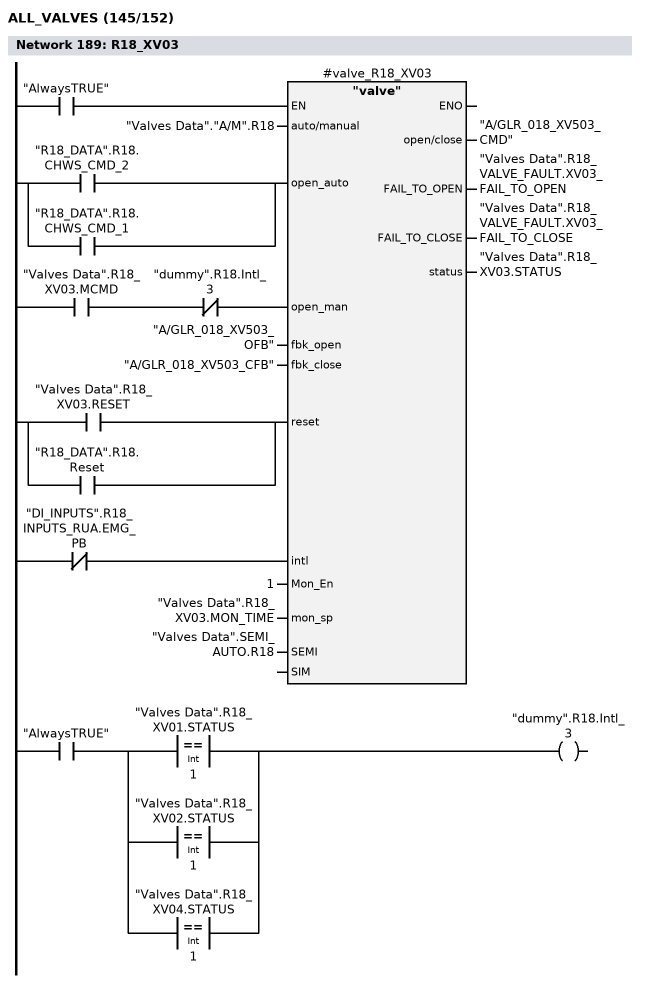
   RUNG wire#powerrail
      Contact( "AlwaysTRUE" )
      #valve_R18_XV03(open_auto := wire#w1, open_man := wire#w2, reset := wire#w3, intl := wire#w4, "auto/manual" := "Valves Data"."A/M".R18, fbk_open := "A/GLR_018_XV503_OFB", fbk_close := "A/GLR_018_XV503_CFB", Mon_En := 1, mon_sp := "Valves Data".R18_XV03.MON_TIME, SEMI := "Valves Data".SEMI_AUTO.R18, SIM :=, "open/close" => "A/GLR_018_XV503_CMD", FAIL_TO_OPEN => "Valves Data".R18_VALVE_FAULT.XV03_FAIL_TO_OPEN, FAIL_TO_CLOSE => "Valves Data".R18_VALVE_FAULT.XV03_FAIL_TO_CLOSE, status => "Valves Data".R18_XV03.STATUS)
   END_RUNG
   RUNG wire#powerrail
      Contact( "R18_DATA".R18.CHWS_CMD_2 )
   END_RUNG wire#w1
   RUNG wire#powerrail
      Contact( "R18_DATA".R18.CHWS_CMD_1 )
   END_RUNG wire#w1
   RUNG wire#powerrail
      Contact( "Valves Data".R18_XV03.MCMD )
      I_Contact( "dummy".R18.Intl_3 )
   END_RUNG wire#w2
   RUNG wire#powerrail
      Contact( "Valves Data".R18_XV03.RESET )
   END_RUNG wire#w3
   RUNG wire#powerrail
      Contact( "R18_DATA".R18.Reset )
   END_RUNG wire#w3
   RUNG wire#powerrail
      I_Contact( "DI_INPUTS".R18_INPUTS_RUA.EMG_PB )
   END_RUNG wire#w4
   RUNG wire#powerrail
      Contact( "AlwaysTRUE" )
      wire#w5
      { S7_Templates := "SrcType := Int" } EQ_Contact(in1 := "Valves Data".R18_XV01.STATUS, in2 := 1)
      wire#w6
      Coil( "dummy".R18.Intl_3 )
   END_RUNG
   RUNG wire#w5
      { S7_Templates := "SrcType := Int" } EQ_Contact(in1 := "Valves Data".R18_XV02.STATUS, in2 := 1)
   END_RUNG wire#w6
   RUNG wire#w5
      { S7_Templates := "SrcType := Int" } EQ_Contact(in1 := "Valves Data".R18_XV04.STATUS, in2 := 1)
   END_RUNG wire#w6
   // the same network as SCL:
   IF "AlwaysTRUE" THEN
       #valve_R18_XV03("auto/manual" := "Valves Data"."A/M".R18,   // "valve"
                       open_auto := "R18_DATA".R18.CHWS_CMD_2 OR "R18_DATA".R18.CHWS_CMD_1,
                       open_man := "Valves Data".R18_XV03.MCMD AND NOT "dummy".R18.Intl_3,
                       fbk_open := "A/GLR_018_XV503_OFB",
                       fbk_close := "A/GLR_018_XV503_CFB",
                       reset := "Valves Data".R18_XV03.RESET OR "R18_DATA".R18.Reset,
                       intl := NOT "DI_INPUTS".R18_INPUTS_RUA.EMG_PB,
                       Mon_En := 1,
                       mon_sp := "Valves Data".R18_XV03.MON_TIME,
                       SEMI := "Valves Data".SEMI_AUTO.R18,
                       "open/close" => "A/GLR_018_XV503_CMD",
                       FAIL_TO_OPEN => "Valves Data".R18_VALVE_FAULT.XV03_FAIL_TO_OPEN,
                       FAIL_TO_CLOSE => "Valves Data".R18_VALVE_FAULT.XV03_FAIL_TO_CLOSE,
                       status => "Valves Data".R18_XV03.STATUS);
   END_IF;
   "dummy".R18.Intl_3 := "AlwaysTRUE" AND (("Valves Data".R18_XV01.STATUS = 1) OR ("Valves Data".R18_XV02.STATUS = 1) OR ("Valves Data".R18_XV04.STATUS = 1));
END_REGION

REGION Network 190: R18_XV04
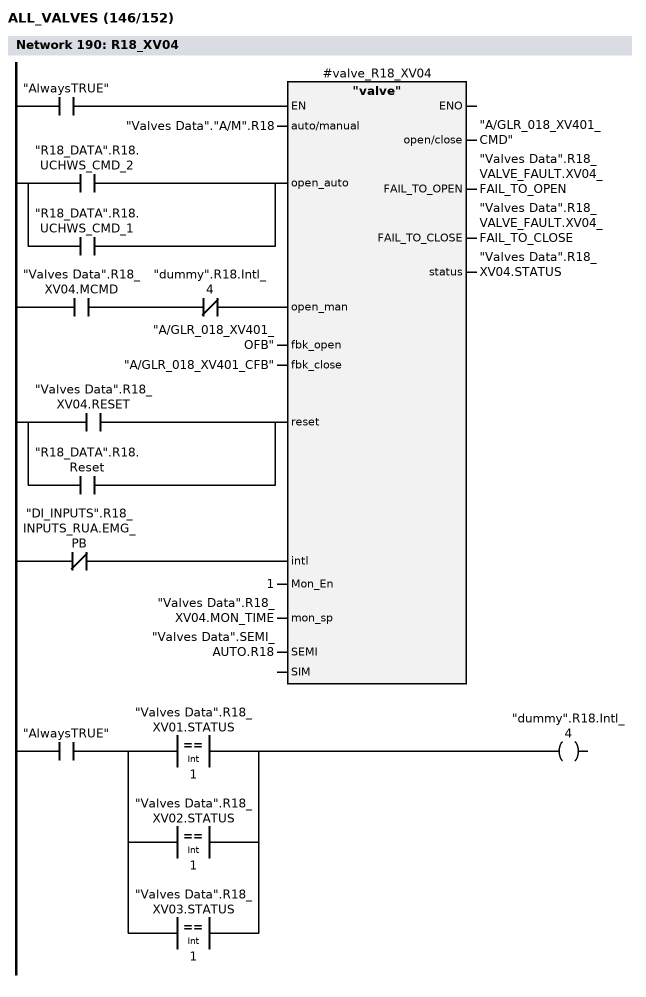
   RUNG wire#powerrail
      Contact( "AlwaysTRUE" )
      #valve_R18_XV04(open_auto := wire#w1, open_man := wire#w2, reset := wire#w3, intl := wire#w4, "auto/manual" := "Valves Data"."A/M".R18, fbk_open := "A/GLR_018_XV401_OFB", fbk_close := "A/GLR_018_XV401_CFB", Mon_En := 1, mon_sp := "Valves Data".R18_XV04.MON_TIME, SEMI := "Valves Data".SEMI_AUTO.R18, SIM :=, "open/close" => "A/GLR_018_XV401_CMD", FAIL_TO_OPEN => "Valves Data".R18_VALVE_FAULT.XV04_FAIL_TO_OPEN, FAIL_TO_CLOSE => "Valves Data".R18_VALVE_FAULT.XV04_FAIL_TO_CLOSE, status => "Valves Data".R18_XV04.STATUS)
   END_RUNG
   RUNG wire#powerrail
      Contact( "R18_DATA".R18.UCHWS_CMD_2 )
   END_RUNG wire#w1
   RUNG wire#powerrail
      Contact( "R18_DATA".R18.UCHWS_CMD_1 )
   END_RUNG wire#w1
   RUNG wire#powerrail
      Contact( "Valves Data".R18_XV04.MCMD )
      I_Contact( "dummy".R18.Intl_4 )
   END_RUNG wire#w2
   RUNG wire#powerrail
      Contact( "Valves Data".R18_XV04.RESET )
   END_RUNG wire#w3
   RUNG wire#powerrail
      Contact( "R18_DATA".R18.Reset )
   END_RUNG wire#w3
   RUNG wire#powerrail
      I_Contact( "DI_INPUTS".R18_INPUTS_RUA.EMG_PB )
   END_RUNG wire#w4
   RUNG wire#powerrail
      Contact( "AlwaysTRUE" )
      wire#w5
      { S7_Templates := "SrcType := Int" } EQ_Contact(in1 := "Valves Data".R18_XV01.STATUS, in2 := 1)
      wire#w6
      Coil( "dummy".R18.Intl_4 )
   END_RUNG
   RUNG wire#w5
      { S7_Templates := "SrcType := Int" } EQ_Contact(in1 := "Valves Data".R18_XV02.STATUS, in2 := 1)
   END_RUNG wire#w6
   RUNG wire#w5
      { S7_Templates := "SrcType := Int" } EQ_Contact(in1 := "Valves Data".R18_XV03.STATUS, in2 := 1)
   END_RUNG wire#w6
   // the same network as SCL:
   IF "AlwaysTRUE" THEN
       #valve_R18_XV04("auto/manual" := "Valves Data"."A/M".R18,   // "valve"
                       open_auto := "R18_DATA".R18.UCHWS_CMD_2 OR "R18_DATA".R18.UCHWS_CMD_1,
                       open_man := "Valves Data".R18_XV04.MCMD AND NOT "dummy".R18.Intl_4,
                       fbk_open := "A/GLR_018_XV401_OFB",
                       fbk_close := "A/GLR_018_XV401_CFB",
                       reset := "Valves Data".R18_XV04.RESET OR "R18_DATA".R18.Reset,
                       intl := NOT "DI_INPUTS".R18_INPUTS_RUA.EMG_PB,
                       Mon_En := 1,
                       mon_sp := "Valves Data".R18_XV04.MON_TIME,
                       SEMI := "Valves Data".SEMI_AUTO.R18,
                       "open/close" => "A/GLR_018_XV401_CMD",
                       FAIL_TO_OPEN => "Valves Data".R18_VALVE_FAULT.XV04_FAIL_TO_OPEN,
                       FAIL_TO_CLOSE => "Valves Data".R18_VALVE_FAULT.XV04_FAIL_TO_CLOSE,
                       status => "Valves Data".R18_XV04.STATUS);
   END_IF;
   "dummy".R18.Intl_4 := "AlwaysTRUE" AND (("Valves Data".R18_XV01.STATUS = 1) OR ("Valves Data".R18_XV02.STATUS = 1) OR ("Valves Data".R18_XV03.STATUS = 1));
END_REGION

REGION Network 191: R18_XV05
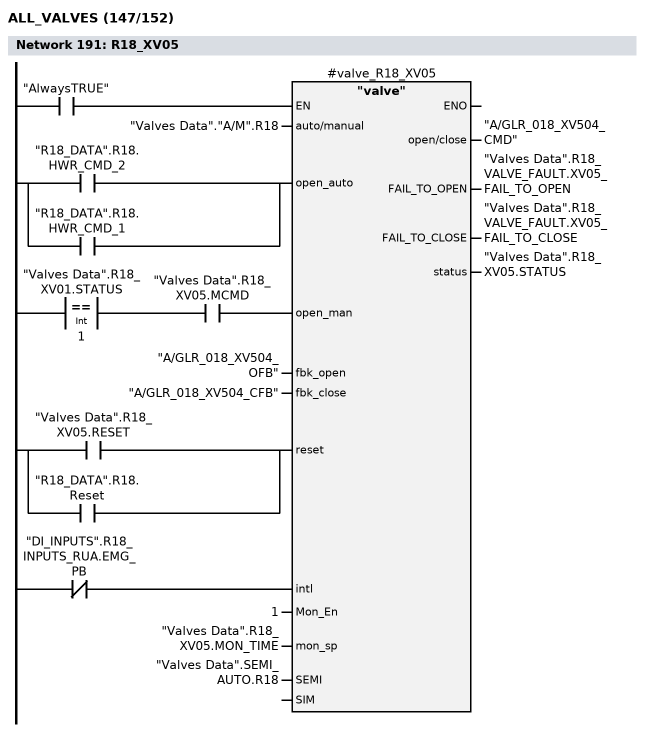
   RUNG wire#powerrail
      Contact( "AlwaysTRUE" )
      #valve_R18_XV05(open_auto := wire#w1, open_man := wire#w2, reset := wire#w3, intl := wire#w4, "auto/manual" := "Valves Data"."A/M".R18, fbk_open := "A/GLR_018_XV504_OFB", fbk_close := "A/GLR_018_XV504_CFB", Mon_En := 1, mon_sp := "Valves Data".R18_XV05.MON_TIME, SEMI := "Valves Data".SEMI_AUTO.R18, SIM :=, "open/close" => "A/GLR_018_XV504_CMD", FAIL_TO_OPEN => "Valves Data".R18_VALVE_FAULT.XV05_FAIL_TO_OPEN, FAIL_TO_CLOSE => "Valves Data".R18_VALVE_FAULT.XV05_FAIL_TO_CLOSE, status => "Valves Data".R18_XV05.STATUS)
   END_RUNG
   RUNG wire#powerrail
      Contact( "R18_DATA".R18.HWR_CMD_2 )
   END_RUNG wire#w1
   RUNG wire#powerrail
      Contact( "R18_DATA".R18.HWR_CMD_1 )
   END_RUNG wire#w1
   RUNG wire#powerrail
      { S7_Templates := "SrcType := Int" } EQ_Contact(in1 := "Valves Data".R18_XV01.STATUS, in2 := 1)
      Contact( "Valves Data".R18_XV05.MCMD )
   END_RUNG wire#w2
   RUNG wire#powerrail
      Contact( "Valves Data".R18_XV05.RESET )
   END_RUNG wire#w3
   RUNG wire#powerrail
      Contact( "R18_DATA".R18.Reset )
   END_RUNG wire#w3
   RUNG wire#powerrail
      I_Contact( "DI_INPUTS".R18_INPUTS_RUA.EMG_PB )
   END_RUNG wire#w4
   // the same network as SCL:
   IF "AlwaysTRUE" THEN
       #valve_R18_XV05("auto/manual" := "Valves Data"."A/M".R18,   // "valve"
                       open_auto := "R18_DATA".R18.HWR_CMD_2 OR "R18_DATA".R18.HWR_CMD_1,
                       open_man := ("Valves Data".R18_XV01.STATUS = 1) AND "Valves Data".R18_XV05.MCMD,
                       fbk_open := "A/GLR_018_XV504_OFB",
                       fbk_close := "A/GLR_018_XV504_CFB",
                       reset := "Valves Data".R18_XV05.RESET OR "R18_DATA".R18.Reset,
                       intl := NOT "DI_INPUTS".R18_INPUTS_RUA.EMG_PB,
                       Mon_En := 1,
                       mon_sp := "Valves Data".R18_XV05.MON_TIME,
                       SEMI := "Valves Data".SEMI_AUTO.R18,
                       "open/close" => "A/GLR_018_XV504_CMD",
                       FAIL_TO_OPEN => "Valves Data".R18_VALVE_FAULT.XV05_FAIL_TO_OPEN,
                       FAIL_TO_CLOSE => "Valves Data".R18_VALVE_FAULT.XV05_FAIL_TO_CLOSE,
                       status => "Valves Data".R18_XV05.STATUS);
   END_IF;
END_REGION

REGION Network 192: R18_XV06
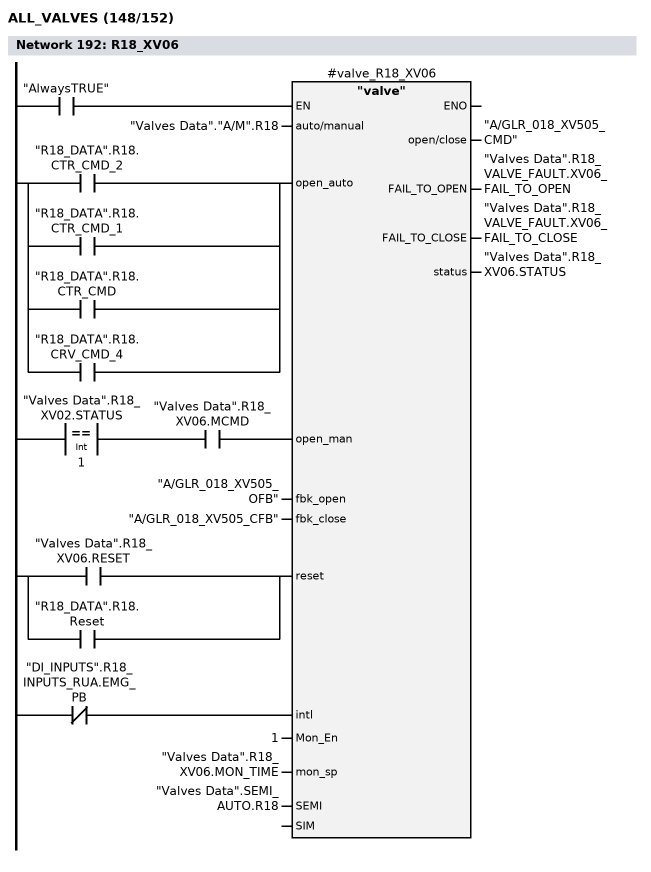
   RUNG wire#powerrail
      Contact( "AlwaysTRUE" )
      #valve_R18_XV06(open_auto := wire#w1, open_man := wire#w2, reset := wire#w3, intl := wire#w4, "auto/manual" := "Valves Data"."A/M".R18, fbk_open := "A/GLR_018_XV505_OFB", fbk_close := "A/GLR_018_XV505_CFB", Mon_En := 1, mon_sp := "Valves Data".R18_XV06.MON_TIME, SEMI := "Valves Data".SEMI_AUTO.R18, SIM :=, "open/close" => "A/GLR_018_XV505_CMD", FAIL_TO_OPEN => "Valves Data".R18_VALVE_FAULT.XV06_FAIL_TO_OPEN, FAIL_TO_CLOSE => "Valves Data".R18_VALVE_FAULT.XV06_FAIL_TO_CLOSE, status => "Valves Data".R18_XV06.STATUS)
   END_RUNG
   RUNG wire#powerrail
      Contact( "R18_DATA".R18.CTR_CMD_2 )
   END_RUNG wire#w1
   RUNG wire#powerrail
      Contact( "R18_DATA".R18.CTR_CMD_1 )
   END_RUNG wire#w1
   RUNG wire#powerrail
      Contact( "R18_DATA".R18.CTR_CMD )
   END_RUNG wire#w1
   RUNG wire#powerrail
      Contact( "R18_DATA".R18.CRV_CMD_4 )
   END_RUNG wire#w1
   RUNG wire#powerrail
      { S7_Templates := "SrcType := Int" } EQ_Contact(in1 := "Valves Data".R18_XV02.STATUS, in2 := 1)
      Contact( "Valves Data".R18_XV06.MCMD )
   END_RUNG wire#w2
   RUNG wire#powerrail
      Contact( "Valves Data".R18_XV06.RESET )
   END_RUNG wire#w3
   RUNG wire#powerrail
      Contact( "R18_DATA".R18.Reset )
   END_RUNG wire#w3
   RUNG wire#powerrail
      I_Contact( "DI_INPUTS".R18_INPUTS_RUA.EMG_PB )
   END_RUNG wire#w4
   // the same network as SCL:
   IF "AlwaysTRUE" THEN
       #valve_R18_XV06("auto/manual" := "Valves Data"."A/M".R18,   // "valve"
                       open_auto := "R18_DATA".R18.CTR_CMD_2 OR "R18_DATA".R18.CTR_CMD_1 OR "R18_DATA".R18.CTR_CMD OR "R18_DATA".R18.CRV_CMD_4,
                       open_man := ("Valves Data".R18_XV02.STATUS = 1) AND "Valves Data".R18_XV06.MCMD,
                       fbk_open := "A/GLR_018_XV505_OFB",
                       fbk_close := "A/GLR_018_XV505_CFB",
                       reset := "Valves Data".R18_XV06.RESET OR "R18_DATA".R18.Reset,
                       intl := NOT "DI_INPUTS".R18_INPUTS_RUA.EMG_PB,
                       Mon_En := 1,
                       mon_sp := "Valves Data".R18_XV06.MON_TIME,
                       SEMI := "Valves Data".SEMI_AUTO.R18,
                       "open/close" => "A/GLR_018_XV505_CMD",
                       FAIL_TO_OPEN => "Valves Data".R18_VALVE_FAULT.XV06_FAIL_TO_OPEN,
                       FAIL_TO_CLOSE => "Valves Data".R18_VALVE_FAULT.XV06_FAIL_TO_CLOSE,
                       status => "Valves Data".R18_XV06.STATUS);
   END_IF;
END_REGION

REGION Network 193: R18_XV07
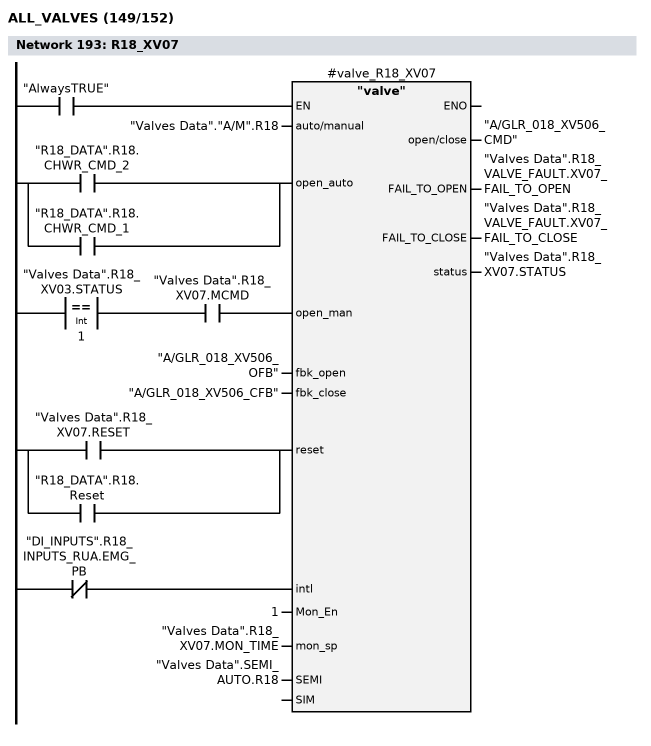
   RUNG wire#powerrail
      Contact( "AlwaysTRUE" )
      #valve_R18_XV07(open_auto := wire#w1, open_man := wire#w2, reset := wire#w3, intl := wire#w4, "auto/manual" := "Valves Data"."A/M".R18, fbk_open := "A/GLR_018_XV506_OFB", fbk_close := "A/GLR_018_XV506_CFB", Mon_En := 1, mon_sp := "Valves Data".R18_XV07.MON_TIME, SEMI := "Valves Data".SEMI_AUTO.R18, SIM :=, "open/close" => "A/GLR_018_XV506_CMD", FAIL_TO_OPEN => "Valves Data".R18_VALVE_FAULT.XV07_FAIL_TO_OPEN, FAIL_TO_CLOSE => "Valves Data".R18_VALVE_FAULT.XV07_FAIL_TO_CLOSE, status => "Valves Data".R18_XV07.STATUS)
   END_RUNG
   RUNG wire#powerrail
      Contact( "R18_DATA".R18.CHWR_CMD_2 )
   END_RUNG wire#w1
   RUNG wire#powerrail
      Contact( "R18_DATA".R18.CHWR_CMD_1 )
   END_RUNG wire#w1
   RUNG wire#powerrail
      { S7_Templates := "SrcType := Int" } EQ_Contact(in1 := "Valves Data".R18_XV03.STATUS, in2 := 1)
      Contact( "Valves Data".R18_XV07.MCMD )
   END_RUNG wire#w2
   RUNG wire#powerrail
      Contact( "Valves Data".R18_XV07.RESET )
   END_RUNG wire#w3
   RUNG wire#powerrail
      Contact( "R18_DATA".R18.Reset )
   END_RUNG wire#w3
   RUNG wire#powerrail
      I_Contact( "DI_INPUTS".R18_INPUTS_RUA.EMG_PB )
   END_RUNG wire#w4
   // the same network as SCL:
   IF "AlwaysTRUE" THEN
       #valve_R18_XV07("auto/manual" := "Valves Data"."A/M".R18,   // "valve"
                       open_auto := "R18_DATA".R18.CHWR_CMD_2 OR "R18_DATA".R18.CHWR_CMD_1,
                       open_man := ("Valves Data".R18_XV03.STATUS = 1) AND "Valves Data".R18_XV07.MCMD,
                       fbk_open := "A/GLR_018_XV506_OFB",
                       fbk_close := "A/GLR_018_XV506_CFB",
                       reset := "Valves Data".R18_XV07.RESET OR "R18_DATA".R18.Reset,
                       intl := NOT "DI_INPUTS".R18_INPUTS_RUA.EMG_PB,
                       Mon_En := 1,
                       mon_sp := "Valves Data".R18_XV07.MON_TIME,
                       SEMI := "Valves Data".SEMI_AUTO.R18,
                       "open/close" => "A/GLR_018_XV506_CMD",
                       FAIL_TO_OPEN => "Valves Data".R18_VALVE_FAULT.XV07_FAIL_TO_OPEN,
                       FAIL_TO_CLOSE => "Valves Data".R18_VALVE_FAULT.XV07_FAIL_TO_CLOSE,
                       status => "Valves Data".R18_XV07.STATUS);
   END_IF;
END_REGION

REGION Network 194: R18_XV08
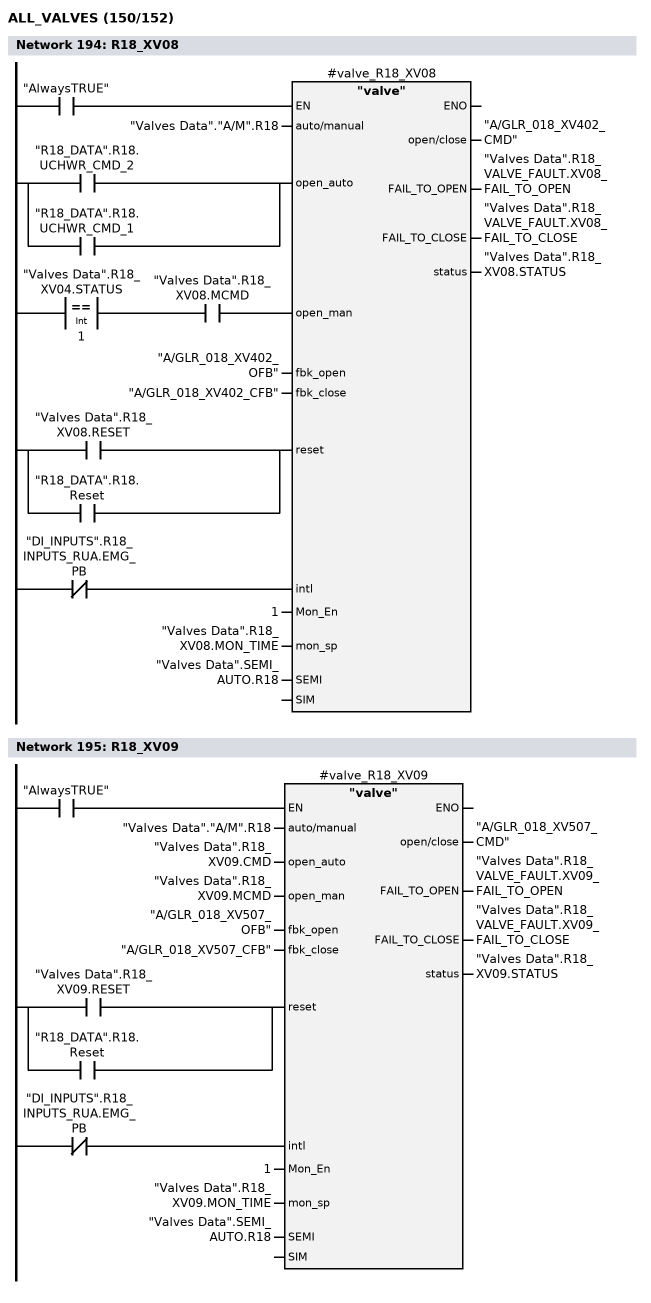
   RUNG wire#powerrail
      Contact( "AlwaysTRUE" )
      #valve_R18_XV08(open_auto := wire#w1, open_man := wire#w2, reset := wire#w3, intl := wire#w4, "auto/manual" := "Valves Data"."A/M".R18, fbk_open := "A/GLR_018_XV402_OFB", fbk_close := "A/GLR_018_XV402_CFB", Mon_En := 1, mon_sp := "Valves Data".R18_XV08.MON_TIME, SEMI := "Valves Data".SEMI_AUTO.R18, SIM :=, "open/close" => "A/GLR_018_XV402_CMD", FAIL_TO_OPEN => "Valves Data".R18_VALVE_FAULT.XV08_FAIL_TO_OPEN, FAIL_TO_CLOSE => "Valves Data".R18_VALVE_FAULT.XV08_FAIL_TO_CLOSE, status => "Valves Data".R18_XV08.STATUS)
   END_RUNG
   RUNG wire#powerrail
      Contact( "R18_DATA".R18.UCHWR_CMD_2 )
   END_RUNG wire#w1
   RUNG wire#powerrail
      Contact( "R18_DATA".R18.UCHWR_CMD_1 )
   END_RUNG wire#w1
   RUNG wire#powerrail
      { S7_Templates := "SrcType := Int" } EQ_Contact(in1 := "Valves Data".R18_XV04.STATUS, in2 := 1)
      Contact( "Valves Data".R18_XV08.MCMD )
   END_RUNG wire#w2
   RUNG wire#powerrail
      Contact( "Valves Data".R18_XV08.RESET )
   END_RUNG wire#w3
   RUNG wire#powerrail
      Contact( "R18_DATA".R18.Reset )
   END_RUNG wire#w3
   RUNG wire#powerrail
      I_Contact( "DI_INPUTS".R18_INPUTS_RUA.EMG_PB )
   END_RUNG wire#w4
   // the same network as SCL:
   IF "AlwaysTRUE" THEN
       #valve_R18_XV08("auto/manual" := "Valves Data"."A/M".R18,   // "valve"
                       open_auto := "R18_DATA".R18.UCHWR_CMD_2 OR "R18_DATA".R18.UCHWR_CMD_1,
                       open_man := ("Valves Data".R18_XV04.STATUS = 1) AND "Valves Data".R18_XV08.MCMD,
                       fbk_open := "A/GLR_018_XV402_OFB",
                       fbk_close := "A/GLR_018_XV402_CFB",
                       reset := "Valves Data".R18_XV08.RESET OR "R18_DATA".R18.Reset,
                       intl := NOT "DI_INPUTS".R18_INPUTS_RUA.EMG_PB,
                       Mon_En := 1,
                       mon_sp := "Valves Data".R18_XV08.MON_TIME,
                       SEMI := "Valves Data".SEMI_AUTO.R18,
                       "open/close" => "A/GLR_018_XV402_CMD",
                       FAIL_TO_OPEN => "Valves Data".R18_VALVE_FAULT.XV08_FAIL_TO_OPEN,
                       FAIL_TO_CLOSE => "Valves Data".R18_VALVE_FAULT.XV08_FAIL_TO_CLOSE,
                       status => "Valves Data".R18_XV08.STATUS);
   END_IF;
END_REGION

REGION Network 195: R18_XV09
   RUNG wire#powerrail
      Contact( "AlwaysTRUE" )
      #valve_R18_XV09(reset := wire#w1, intl := wire#w2, "auto/manual" := "Valves Data"."A/M".R18, open_auto := "Valves Data".R18_XV09.CMD, open_man := "Valves Data".R18_XV09.MCMD, fbk_open := "A/GLR_018_XV507_OFB", fbk_close := "A/GLR_018_XV507_CFB", Mon_En := 1, mon_sp := "Valves Data".R18_XV09.MON_TIME, SEMI := "Valves Data".SEMI_AUTO.R18, SIM :=, "open/close" => "A/GLR_018_XV507_CMD", FAIL_TO_OPEN => "Valves Data".R18_VALVE_FAULT.XV09_FAIL_TO_OPEN, FAIL_TO_CLOSE => "Valves Data".R18_VALVE_FAULT.XV09_FAIL_TO_CLOSE, status => "Valves Data".R18_XV09.STATUS)
   END_RUNG
   RUNG wire#powerrail
      Contact( "Valves Data".R18_XV09.RESET )
   END_RUNG wire#w1
   RUNG wire#powerrail
      Contact( "R18_DATA".R18.Reset )
   END_RUNG wire#w1
   RUNG wire#powerrail
      I_Contact( "DI_INPUTS".R18_INPUTS_RUA.EMG_PB )
   END_RUNG wire#w2
   // the same network as SCL:
   IF "AlwaysTRUE" THEN
       #valve_R18_XV09("auto/manual" := "Valves Data"."A/M".R18,   // "valve"
                       open_auto := "Valves Data".R18_XV09.CMD,
                       open_man := "Valves Data".R18_XV09.MCMD,
                       fbk_open := "A/GLR_018_XV507_OFB",
                       fbk_close := "A/GLR_018_XV507_CFB",
                       reset := "Valves Data".R18_XV09.RESET OR "R18_DATA".R18.Reset,
                       intl := NOT "DI_INPUTS".R18_INPUTS_RUA.EMG_PB,
                       Mon_En := 1,
                       mon_sp := "Valves Data".R18_XV09.MON_TIME,
                       SEMI := "Valves Data".SEMI_AUTO.R18,
                       "open/close" => "A/GLR_018_XV507_CMD",
                       FAIL_TO_OPEN => "Valves Data".R18_VALVE_FAULT.XV09_FAIL_TO_OPEN,
                       FAIL_TO_CLOSE => "Valves Data".R18_VALVE_FAULT.XV09_FAIL_TO_CLOSE,
                       status => "Valves Data".R18_XV09.STATUS);
   END_IF;
END_REGION

REGION Network 196: R18_XV10
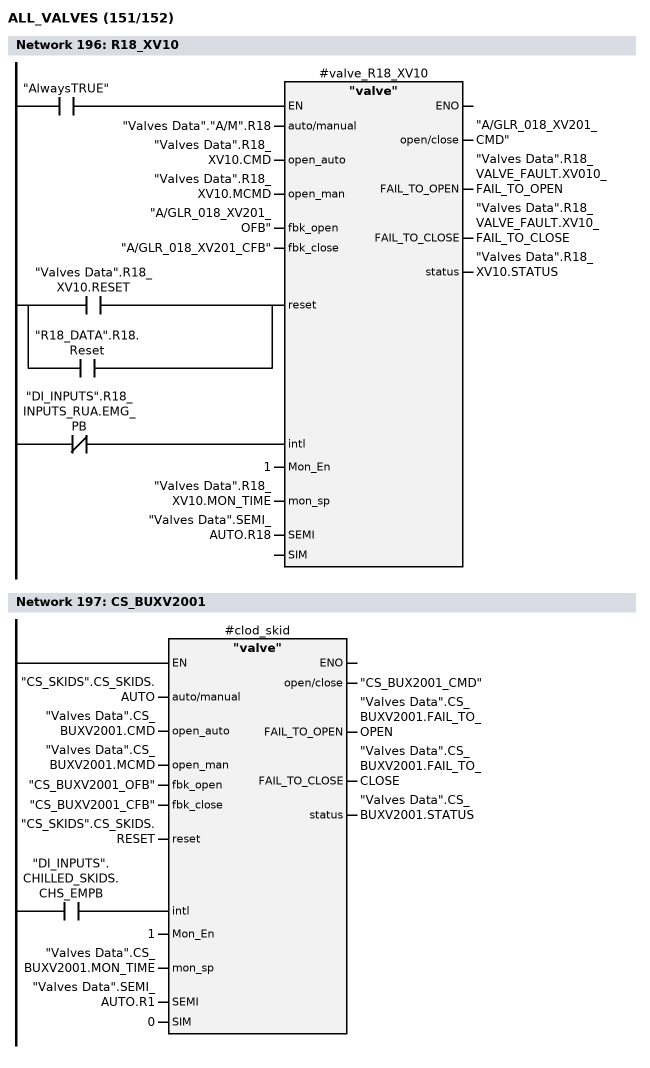
   RUNG wire#powerrail
      Contact( "AlwaysTRUE" )
      #valve_R18_XV10(reset := wire#w1, intl := wire#w2, "auto/manual" := "Valves Data"."A/M".R18, open_auto := "Valves Data".R18_XV10.CMD, open_man := "Valves Data".R18_XV10.MCMD, fbk_open := "A/GLR_018_XV201_OFB", fbk_close := "A/GLR_018_XV201_CFB", Mon_En := 1, mon_sp := "Valves Data".R18_XV10.MON_TIME, SEMI := "Valves Data".SEMI_AUTO.R18, SIM :=, "open/close" => "A/GLR_018_XV201_CMD", FAIL_TO_OPEN => "Valves Data".R18_VALVE_FAULT.XV010_FAIL_TO_OPEN, FAIL_TO_CLOSE => "Valves Data".R18_VALVE_FAULT.XV10_FAIL_TO_CLOSE, status => "Valves Data".R18_XV10.STATUS)
   END_RUNG
   RUNG wire#powerrail
      Contact( "Valves Data".R18_XV10.RESET )
   END_RUNG wire#w1
   RUNG wire#powerrail
      Contact( "R18_DATA".R18.Reset )
   END_RUNG wire#w1
   RUNG wire#powerrail
      I_Contact( "DI_INPUTS".R18_INPUTS_RUA.EMG_PB )
   END_RUNG wire#w2
   // the same network as SCL:
   IF "AlwaysTRUE" THEN
       #valve_R18_XV10("auto/manual" := "Valves Data"."A/M".R18,   // "valve"
                       open_auto := "Valves Data".R18_XV10.CMD,
                       open_man := "Valves Data".R18_XV10.MCMD,
                       fbk_open := "A/GLR_018_XV201_OFB",
                       fbk_close := "A/GLR_018_XV201_CFB",
                       reset := "Valves Data".R18_XV10.RESET OR "R18_DATA".R18.Reset,
                       intl := NOT "DI_INPUTS".R18_INPUTS_RUA.EMG_PB,
                       Mon_En := 1,
                       mon_sp := "Valves Data".R18_XV10.MON_TIME,
                       SEMI := "Valves Data".SEMI_AUTO.R18,
                       "open/close" => "A/GLR_018_XV201_CMD",
                       FAIL_TO_OPEN => "Valves Data".R18_VALVE_FAULT.XV010_FAIL_TO_OPEN,
                       FAIL_TO_CLOSE => "Valves Data".R18_VALVE_FAULT.XV10_FAIL_TO_CLOSE,
                       status => "Valves Data".R18_XV10.STATUS);
   END_IF;
END_REGION

REGION Network 197: CS_BUXV2001
   RUNG wire#powerrail
      #clod_skid(intl := wire#w1, "auto/manual" := "CS_SKIDS".CS_SKIDS.AUTO, open_auto := "Valves Data".CS_BUXV2001.CMD, open_man := "Valves Data".CS_BUXV2001.MCMD, fbk_open := "CS_BUXV2001_OFB", fbk_close := "CS_BUXV2001_CFB", reset := "CS_SKIDS".CS_SKIDS.RESET, Mon_En := 1, mon_sp := "Valves Data".CS_BUXV2001.MON_TIME, SEMI := "Valves Data".SEMI_AUTO.R1, SIM := 0, "open/close" => "CS_BUX2001_CMD", FAIL_TO_OPEN => "Valves Data".CS_BUXV2001.FAIL_TO_OPEN, FAIL_TO_CLOSE => "Valves Data".CS_BUXV2001.FAIL_TO_CLOSE, status => "Valves Data".CS_BUXV2001.STATUS)
   END_RUNG
   RUNG wire#powerrail
      Contact( "DI_INPUTS".CHILLED_SKIDS.CHS_EMPB )
   END_RUNG wire#w1
   // the same network as SCL:
   #clod_skid("auto/manual" := "CS_SKIDS".CS_SKIDS.AUTO,   // "valve"
              open_auto := "Valves Data".CS_BUXV2001.CMD,
              open_man := "Valves Data".CS_BUXV2001.MCMD,
              fbk_open := "CS_BUXV2001_OFB",
              fbk_close := "CS_BUXV2001_CFB",
              reset := "CS_SKIDS".CS_SKIDS.RESET,
              intl := "DI_INPUTS".CHILLED_SKIDS.CHS_EMPB,
              Mon_En := 1,
              mon_sp := "Valves Data".CS_BUXV2001.MON_TIME,
              SEMI := "Valves Data".SEMI_AUTO.R1,
              SIM := 0,
              "open/close" => "CS_BUX2001_CMD",
              FAIL_TO_OPEN => "Valves Data".CS_BUXV2001.FAIL_TO_OPEN,
              FAIL_TO_CLOSE => "Valves Data".CS_BUXV2001.FAIL_TO_CLOSE,
              status => "Valves Data".CS_BUXV2001.STATUS);
END_REGION

REGION Network 198: UCHS_BUXV1501
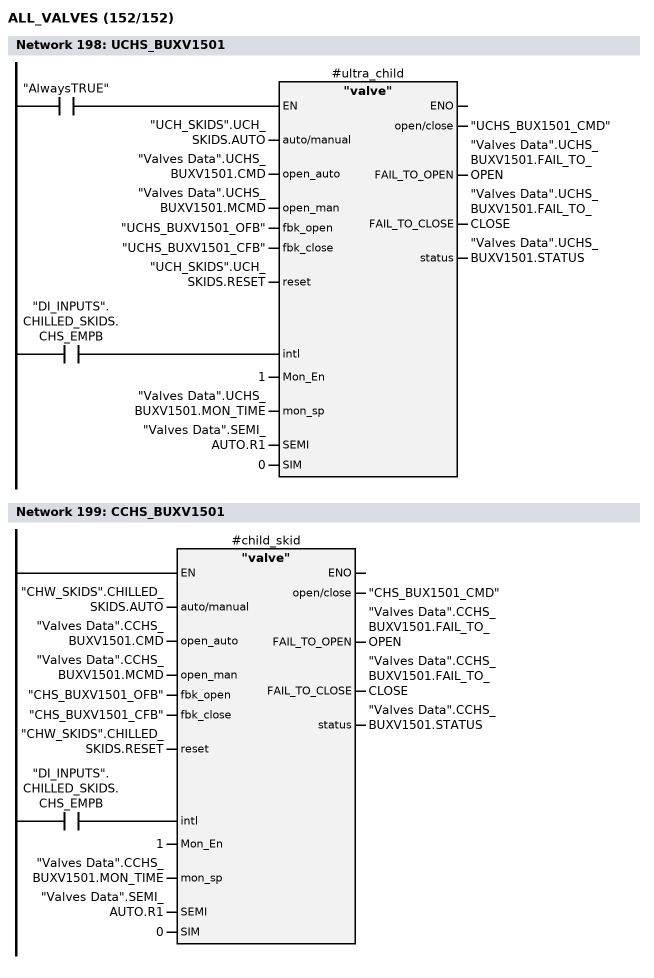
   RUNG wire#powerrail
      Contact( "AlwaysTRUE" )
      #ultra_child(intl := wire#w1, "auto/manual" := "UCH_SKIDS".UCH_SKIDS.AUTO, open_auto := "Valves Data".UCHS_BUXV1501.CMD, open_man := "Valves Data".UCHS_BUXV1501.MCMD, fbk_open := "UCHS_BUXV1501_OFB", fbk_close := "UCHS_BUXV1501_CFB", reset := "UCH_SKIDS".UCH_SKIDS.RESET, Mon_En := 1, mon_sp := "Valves Data".UCHS_BUXV1501.MON_TIME, SEMI := "Valves Data".SEMI_AUTO.R1, SIM := 0, "open/close" => "UCHS_BUX1501_CMD", FAIL_TO_OPEN => "Valves Data".UCHS_BUXV1501.FAIL_TO_OPEN, FAIL_TO_CLOSE => "Valves Data".UCHS_BUXV1501.FAIL_TO_CLOSE, status => "Valves Data".UCHS_BUXV1501.STATUS)
   END_RUNG
   RUNG wire#powerrail
      Contact( "DI_INPUTS".CHILLED_SKIDS.CHS_EMPB )
   END_RUNG wire#w1
   // the same network as SCL:
   IF "AlwaysTRUE" THEN
       #ultra_child("auto/manual" := "UCH_SKIDS".UCH_SKIDS.AUTO,   // "valve"
                    open_auto := "Valves Data".UCHS_BUXV1501.CMD,
                    open_man := "Valves Data".UCHS_BUXV1501.MCMD,
                    fbk_open := "UCHS_BUXV1501_OFB",
                    fbk_close := "UCHS_BUXV1501_CFB",
                    reset := "UCH_SKIDS".UCH_SKIDS.RESET,
                    intl := "DI_INPUTS".CHILLED_SKIDS.CHS_EMPB,
                    Mon_En := 1,
                    mon_sp := "Valves Data".UCHS_BUXV1501.MON_TIME,
                    SEMI := "Valves Data".SEMI_AUTO.R1,
                    SIM := 0,
                    "open/close" => "UCHS_BUX1501_CMD",
                    FAIL_TO_OPEN => "Valves Data".UCHS_BUXV1501.FAIL_TO_OPEN,
                    FAIL_TO_CLOSE => "Valves Data".UCHS_BUXV1501.FAIL_TO_CLOSE,
                    status => "Valves Data".UCHS_BUXV1501.STATUS);
   END_IF;
END_REGION

REGION Network 199: CCHS_BUXV1501
   RUNG wire#powerrail
      #child_skid(intl := wire#w1, "auto/manual" := "CHW_SKIDS".CHILLED_SKIDS.AUTO, open_auto := "Valves Data".CCHS_BUXV1501.CMD, open_man := "Valves Data".CCHS_BUXV1501.MCMD, fbk_open := "CHS_BUXV1501_OFB", fbk_close := "CHS_BUXV1501_CFB", reset := "CHW_SKIDS".CHILLED_SKIDS.RESET, Mon_En := 1, mon_sp := "Valves Data".CCHS_BUXV1501.MON_TIME, SEMI := "Valves Data".SEMI_AUTO.R1, SIM := 0, "open/close" => "CHS_BUX1501_CMD", FAIL_TO_OPEN => "Valves Data".CCHS_BUXV1501.FAIL_TO_OPEN, FAIL_TO_CLOSE => "Valves Data".CCHS_BUXV1501.FAIL_TO_CLOSE, status => "Valves Data".CCHS_BUXV1501.STATUS)
   END_RUNG
   RUNG wire#powerrail
      Contact( "DI_INPUTS".CHILLED_SKIDS.CHS_EMPB )
   END_RUNG wire#w1
   // the same network as SCL:
   #child_skid("auto/manual" := "CHW_SKIDS".CHILLED_SKIDS.AUTO,   // "valve"
               open_auto := "Valves Data".CCHS_BUXV1501.CMD,
               open_man := "Valves Data".CCHS_BUXV1501.MCMD,
               fbk_open := "CHS_BUXV1501_OFB",
               fbk_close := "CHS_BUXV1501_CFB",
               reset := "CHW_SKIDS".CHILLED_SKIDS.RESET,
               intl := "DI_INPUTS".CHILLED_SKIDS.CHS_EMPB,
               Mon_En := 1,
               mon_sp := "Valves Data".CCHS_BUXV1501.MON_TIME,
               SEMI := "Valves Data".SEMI_AUTO.R1,
               SIM := 0,
               "open/close" => "CHS_BUX1501_CMD",
               FAIL_TO_OPEN => "Valves Data".CCHS_BUXV1501.FAIL_TO_OPEN,
               FAIL_TO_CLOSE => "Valves Data".CCHS_BUXV1501.FAIL_TO_CLOSE,
               status => "Valves Data".CCHS_BUXV1501.STATUS);
END_REGION
END_FUNCTION_BLOCK
